(* Logix 5000 project; controller R400_500_XLS vendor 1 type 14 code 216 rev 31.11; software revision 31.01; part 3 of 32 *)
(* tags used below, declared in another part *)
   Alarm : SINT;   // Wait 3 seconds
   Ashutdown : SINT;   // Not Used
   CURRENT_CYCLE : DINT;
   CycleUsageArraySize : DINT;   // Size of the Cycle Usage Array
   CycleUsageDefaultUserName : STRING;   // Default User Name
   CycleUsageDefaultValue : UDT_CYCLE_USAGE;
   CycleUsageFirstEmptyIndex : DINT;   // Cycle Usage Array First Empty Index
   CycleUsageIterator : DINT;
   CycleUsagePrintoutCycleStartedCount : STRING;
   CycleUsagePrintoutHeader : STRING;
   CycleUsagePrintoutMessage : STRING;
   CycleUsagePrintoutSeparator : STRING;
   CycleUsageSearchCurrentUser : BOOL;
   CycleUsageSearchFirstEmptyIndex : BOOL;
   DESCALER : SINT;
   DRYING : DINT;   // Drying id number
   DRYING_HEAT_SENSITIVE_SEL : DINT;   // Drying heat sensitive
   DRYING_MODE_SEL : DINT;   // Drying mode selector index
   DRYING_TEMP_C_SEL : DINT;   // Drying temperature index
   DRYING_TEMP_F_SEL : DINT;   // Drying temperature index
   DRYING_TEMP_HIGH : REAL;   // Smart drying high temperature set point
   DRYING_TEMP_LOW : REAL;   // Smart drying low temperature set point
   DRYING_TEMP_STANDARD_LOW : REAL;   // Regular drying low temperature set point
   DRYING_TIME_LONG : DINT;   // Smart drying time for heat sensitive mode (in minute)
   DRYING_TIME_MIN_NUM : DINT;   // Drying time (minutes) numeric input index
   DRYING_TIME_SEC_NUM : DINT;   // Drying time (seconds) numeric input index
   DRYING_TIME_SHORT : DINT;   // Smart drying time for heat regular mode (in minute)
   ENVIRO_CARE : SINT;
   EXTRA_CARE : SINT;
   FINALRINSE_1 : DINT;   // Final rinse 1 id number
   FINALRINSE_2 : DINT;   // Final rinse 2 id number
   FINALRINSE_3 : DINT;   // Final rinse 3 id number
   FINALRINSE_4 : DINT;   // Final rinse 4 id number
   FINALRINSE_5 : DINT;   // Final rinse 5 id number
   FINALRINSE_6 : DINT;   // Final rinse 6 id number
   FINALRINSE_7 : DINT;   // Final rinse 7 id number
   FINALRINSE_8 : DINT;   // Final rinse 8 id number
   FINALRINSE_9 : DINT;   // Final rinse 9 id number
   FRINSE_COND_SET_POINT_NUM : DINT;   // Final rinse conductivity set point numeric input index
   FRINSE_DRAIN_SEL : DINT;   // Final rinse drained selector's index
   FRINSE_HEATING_SEL : DINT;   // Final rinse heating selector's index
   FRINSE_MIN_NUMBER_NUM : DINT;   // Final rinse minimum number of final rinse numeric input index
   FRINSE_NUMBER_NUM : DINT;   // Final rinse number of final rinse numeric input index
   FRINSE_RECIRC_SEL : DINT;   // Final rinse recirculated selector's index
   FRINSE_TIME_MIN_NUM : DINT;   // Final rinse time (minutes) numeric input index
   FRINSE_TIME_SEC_NUM : DINT;   // Final rinse time (seconds) numeric input index
   FRINSE_TYPE_SEL : DINT;   // Final rinse type selector's index
   HighLimt : REAL;
   LowLimt : REAL;
   M : DINT[5];   // Memory Bits
   NON_RECIRCULATED_FINAL_RINSE_MINUTES : DINT;   // Number of minutes for the non recirculated final rinse
   NON_RECIRCULATED_FINAL_RINSE_SECONDS : DINT;   // Number of seconds for the non recirculated final rinse
   PLASTIC_CARE : SINT;
   PREWASH_1 : DINT;   // Pre-wash 1 id number
   PREWASH_2 : DINT;   // Pre-wash 2 id number
   PREWASH_3 : DINT;   // Pre-wash 3 id number
   PREWASH_4 : DINT;   // Pre-wash 4 id number
   RINSE_1 : DINT;   // Rinse 1 id number
   RINSE_2 : DINT;   // Rinse 2 id number
   RINSE_3 : DINT;   // Rinse 3 id number
   RINSE_4 : DINT;   // Rinse 4 id number
   RINSE_CARE : SINT;
   Run : DINT;
   sCRLF : STRING;
   Service : DINT[2];   // Unused Service Mode Memory Bit
   sPrntArray : STRING[300];   // Printer String Array
   sSpaceCharacter : STRING;   // Space Character
   STANDARD : SINT;
   String : STRING[50];   // String
   SUMP_HIGH_VOLUME_400 : REAL;   // High sump volume
   SUMP_HIGH_VOLUME_500 : REAL;
   SUMP_LOW_VOLUME_400 : REAL;   // Low sump volume
   SUMP_LOW_VOLUME_500 : REAL;
   Supervisor : DINT;
   Tmr : TIMER[107];
   USER_DEFINED_10 : SINT;
   USER_DEFINED_11 : SINT;
   USER_DEFINED_7 : SINT;
   USER_DEFINED_8 : SINT;
   USER_DEFINED_9 : SINT;
   VENTING : DINT;   // Venting id number
   WASH_1 : DINT;   // Wash 1 id number
   WASH_2 : DINT;   // Wash 2 id number
   WASH_3 : DINT;   // Wash 3 id number
   WASH_4 : DINT;   // Wash 4 id number
   WASH_5 : DINT;   // Wash 5 id number
   WSH41_End_signal : BOOL;   // End of cycle signal
   AlarmTrigger : INT;   // Triggers the alarm screen if different of 0
   bAuditTrailExportButton : BOOL;
   bCSVExportHandshake : BOOL;
   bCycleOrAbortInProcess : BOOL;
   bONSAuditExportTrigger : BOOL;
   bONSAuditTrailEndOfCycle : BOOL;
   bONSBatchReportFileLocation : BOOL;
   bONSManualFileTransfer : BOOL;
   bPushButtonTransferFilesFromSDToUSB : BOOL;
   bTransferFilesFromSDToUSB : BOOL;
   bTransferFilesFromSDToUSBHandshakeLoad : BOOL;
   Current_Screen : DINT;
   CurrentUser : STRING;   // Current User
   CycleUsage : UDT_CYCLE_USAGE[50];
   CycleUsageListSelectedIndex : DINT;   // Current index selected in CycleUsage list
   CycleUsagePrint : BOOL;   // Print Cycle Usage
   CycleUsageResetAllValues : BOOL;   // Reset All Cycle Usage of all user
   CycleUsageResetDate : DINT[7];
   CycleUsageResetSelectedUser : BOOL;   // Reset Cycle Usage for the selected user
   DateTime : DINT[7];
   DISABLE : BOOL;   // Disable bit
   EmailSMSInt : INT[8];   // Email & SMS Notification Integer
   ENABLE : BOOL;   // Enable bit
   FALSE : BOOL;   // Always false bit
   NumInput : UDT_NUMERIC_INPUT[65];   // Numeric input
   PrintIndex : DINT;
   sBatchReportCSVName : STRING;
   sBatchReportFolderPath : STRING;
   Screen_Ctrl : DINT;   // PLC Screen Request
   sCycleCounter : STRING;
   sCycleForFileName : STRING;
   sHyphen : STRING;
   SumpHeatAlmRate : REAL;
   sUnderscore : STRING;
   tAuditTrailRemoteClearHistory : TIMER;
   Tpb : DINT[11];
   TpbImage : DINT[11];
   TRUE : BOOL;   // Always true bit
   udtAuditTrail : UDT_AuditTrail;
   udtCSVDataLogBatchReport : UDT_CSVDataLog;
   udtCSVExport : UDT_CSVExport;
   Unit : Hrdwre;   // Unit Configuration
(* MainProgram, continued *)

ROUTINE Constants   (* structured text *)
// Constant parameters
   // Program constants
   
   // General use constants
   TRUE := 1;				// Permanent, always true bit
   FALSE := 0;				// Permanent, always false bit
   ENABLE := 1;			// Used to ENABLE a bloc function
   DISABLE := 0;			// Used to DISABLE a bloc function
   
   // Sump water volume/level
   SUMP_LOW_VOLUME_400 := 22;        // Sump low water volume in liter
   SUMP_HIGH_VOLUME_400 := 36;       // Sump high water volume in liter
   SUMP_LOW_VOLUME_500 := 28.4;        // Sump low water volume in liter
   SUMP_HIGH_VOLUME_500 := 47.3;       // Sump high water volume in liter
   
   //XLSV10  DGB  2018-09-06 : Adjusted Treatments Constants
   // Treatment constants
   PREWASH_1 := 1;         // Pre-wash 1 id number
   PREWASH_2 := 2;         // Pre-wash 2 id number
   PREWASH_3 := 3;         // Pre-wash 3 id number
   PREWASH_4 := 4;         // Pre-wash 4 id number
   WASH_1 := 5;            // Wash 1 id number
   WASH_2 := 6;            // Wash 2 id number
   WASH_3 := 7;            // Wash 3 id number
   WASH_4 := 8;            // Wash 4 id number
   WASH_5 := 9;            // Wash 5 id number
   RINSE_1 := 10;           // Rinse 1 id number
   RINSE_2 := 11;           // Rinse 2 id number
   RINSE_3 := 12;           // Rinse 3 id number
   RINSE_4 := 13;           // Rinse 4 id number
   FINALRINSE_1 := 14;      // Final rinse 1 id number
   FINALRINSE_2 := 15;     // Final rinse 2 id number
   FINALRINSE_3 := 16;     // Final rinse 3 id number
   FINALRINSE_4 := 17;     // Final rinse 4 id number
   FINALRINSE_5 := 18;     // Final rinse 5 id number
   FINALRINSE_6 := 19;     // Final rinse 6 id number
   FINALRINSE_7 := 20;     // Final rinse 7 id number
   FINALRINSE_8 := 21;     // Final rinse 8 id number
   FINALRINSE_9 := 22;     // Final rinse 9 id number
   DRYING := 23;           // Drying id number
   VENTING := 24;          // Venting id number
   
   // Drying temperature and time
   DRYING_TEMP_LOW := 82.2;   // Smart drying low temperature set point
   DRYING_TEMP_HIGH := 115.6; // Smart drying high temperature set point
   //XLSV10  DGB  2018-09-10 : Changed Regular Low Temperature
   DRYING_TEMP_STANDARD_LOW := 65; // Standard drying high temperature set point
   DRYING_TIME_SHORT := 10;    // Smart drying time for heat regular mode (in minute)
   DRYING_TIME_LONG := 20;     // Smart drying time for heat sensitive mode (in minute)
   
   // Cycle constants
   EXTRA_CARE       := 0;
   ENVIRO_CARE      := 1;
   PLASTIC_CARE     := 2;
   STANDARD         := 3;
   RINSE_CARE       := 4;
   DESCALER         := 5;
   USER_DEFINED_7   := 6;
   USER_DEFINED_8   := 7;
   USER_DEFINED_9   := 8;
   USER_DEFINED_10  := 9;
   USER_DEFINED_11  := 10;
   CURRENT_CYCLE    := 11;
   
   
   // Control lists selectors indexes for the treatement modification
   DRYING_MODE_SEL := 14;
   DRYING_TEMP_C_SEL := 15;
   DRYING_TEMP_F_SEL := 16;
   DRYING_HEAT_SENSITIVE_SEL := 17;
   FRINSE_HEATING_SEL := 18;
   FRINSE_DRAIN_SEL := 19;
   FRINSE_RECIRC_SEL := 20;
   FRINSE_TYPE_SEL := 21;
   
   // Numeric input indexes for the treatement modification
   
   DRYING_TIME_MIN_NUM := 11;
   DRYING_TIME_SEC_NUM := 12;
   FRINSE_TIME_MIN_NUM := 14;
   FRINSE_TIME_SEC_NUM := 15;
   FRINSE_NUMBER_NUM := 16;
   FRINSE_MIN_NUMBER_NUM := 17;
   FRINSE_COND_SET_POINT_NUM := 18;
   
   // Non-recirculated final rinse time
   NON_RECIRCULATED_FINAL_RINSE_MINUTES := 0;
   NON_RECIRCULATED_FINAL_RINSE_SECONDS := 10;
   
   // Sump Heating alarm rate
   SumpHeatAlmRate:= 1.0;
   
   // Pure Water Tank low and High heating limit evaluation steam heated unit
   HighLimt:=0.1;
   LowLimt:=0.0;
   
   
   
   
   
END_ROUTINE

ROUTINE CycleUsage   (* ladder *)
// This Routine contains logic to manage the cycle usage
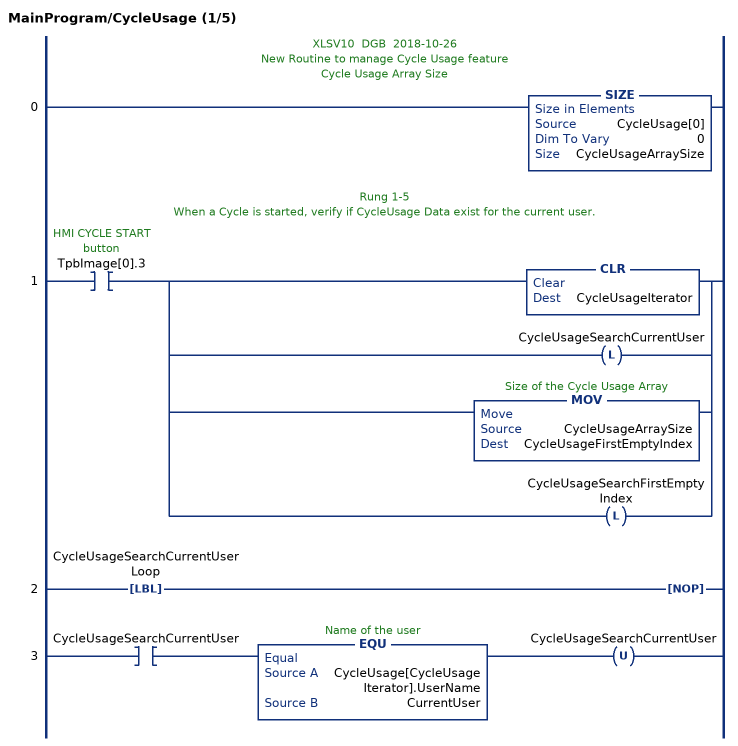
   // XLSV10  DGB  2018-10-26
   //  New Routine to manage Cycle Usage feature
   // Cycle Usage Array Size
   0: SIZE(CycleUsage[0],0,CycleUsageArraySize);
   // Rung 1-5
   // When a Cycle is started, verify if CycleUsage Data exist for the current user.
   1: XIC(TpbImage[0].3)[CLR(CycleUsageIterator) ,OTL(CycleUsageSearchCurrentUser) ,MOV(CycleUsageArraySize,CycleUsageFirstEmptyIndex) ,OTL(CycleUsageSearchFirstEmptyIndex) ];
   2: LBL(CycleUsageSearchCurrentUserLoop)NOP();
   3: XIC(CycleUsageSearchCurrentUser)EQU(CycleUsage[CycleUsageIterator].UserName,CurrentUser)OTU(CycleUsageSearchCurrentUser);
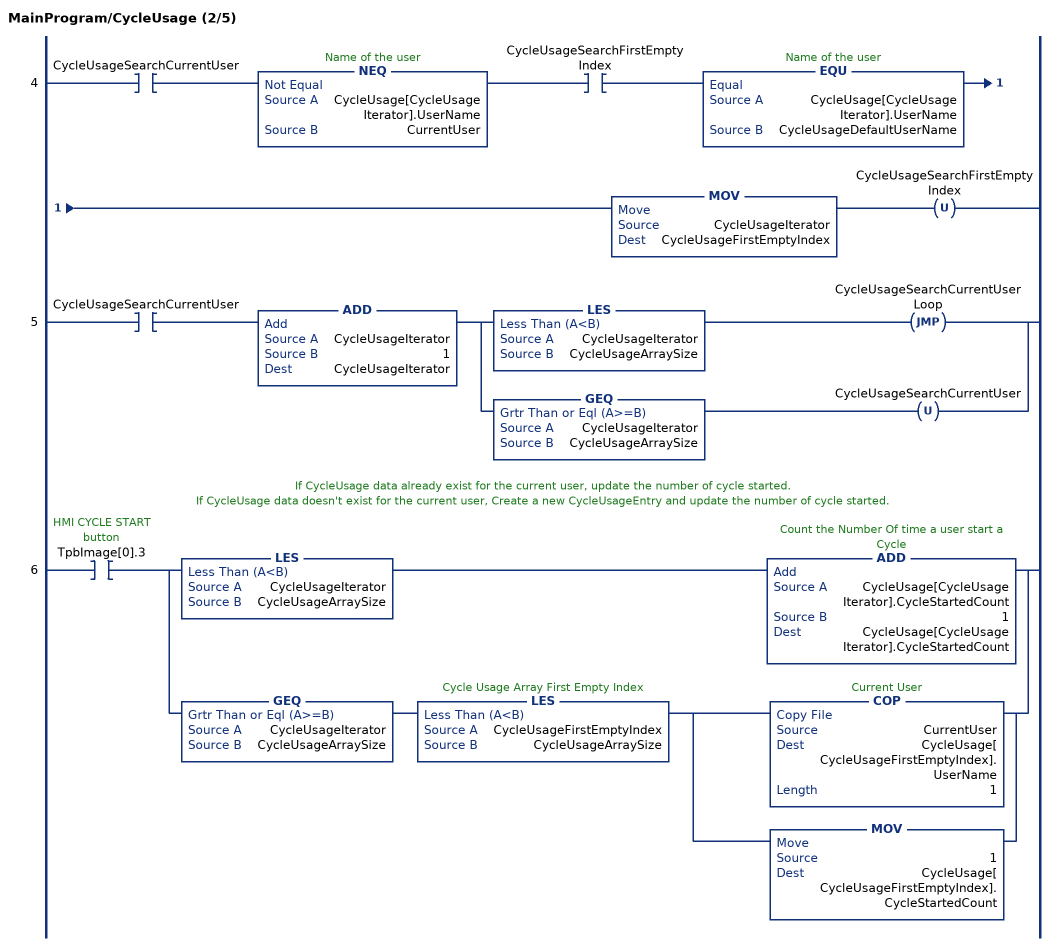
   4: XIC(CycleUsageSearchCurrentUser)NEQ(CycleUsage[CycleUsageIterator].UserName,CurrentUser)XIC(CycleUsageSearchFirstEmptyIndex)EQU(CycleUsage[CycleUsageIterator].UserName,CycleUsageDefaultUserName)MOV(CycleUsageIterator,CycleUsageFirstEmptyIndex)OTU(CycleUsageSearchFirstEmptyIndex);
   5: XIC(CycleUsageSearchCurrentUser)ADD(CycleUsageIterator,1,CycleUsageIterator)[LES(CycleUsageIterator,CycleUsageArraySize) JMP(CycleUsageSearchCurrentUserLoop) ,GEQ(CycleUsageIterator,CycleUsageArraySize) OTU(CycleUsageSearchCurrentUser) ];
   // If CycleUsage data already exist for the current user, update the number of cycle started.
   // If CycleUsage data doesn't exist for the current user, Create a new CycleUsageEntry and update the number of cycle started.
   6: XIC(TpbImage[0].3)[LES(CycleUsageIterator,CycleUsageArraySize) ADD(CycleUsage[CycleUsageIterator].CycleStartedCount,1,CycleUsage[CycleUsageIterator].CycleStartedCount) ,GEQ(CycleUsageIterator,CycleUsageArraySize) LES(CycleUsageFirstEmptyIndex,CycleUsageArraySize) [COP(CurrentUser,CycleUsage[CycleUsageFirstEmptyIndex].UserName,1) ,MOV(1,CycleUsage[CycleUsageFirstEmptyIndex].CycleStartedCount) ] ];
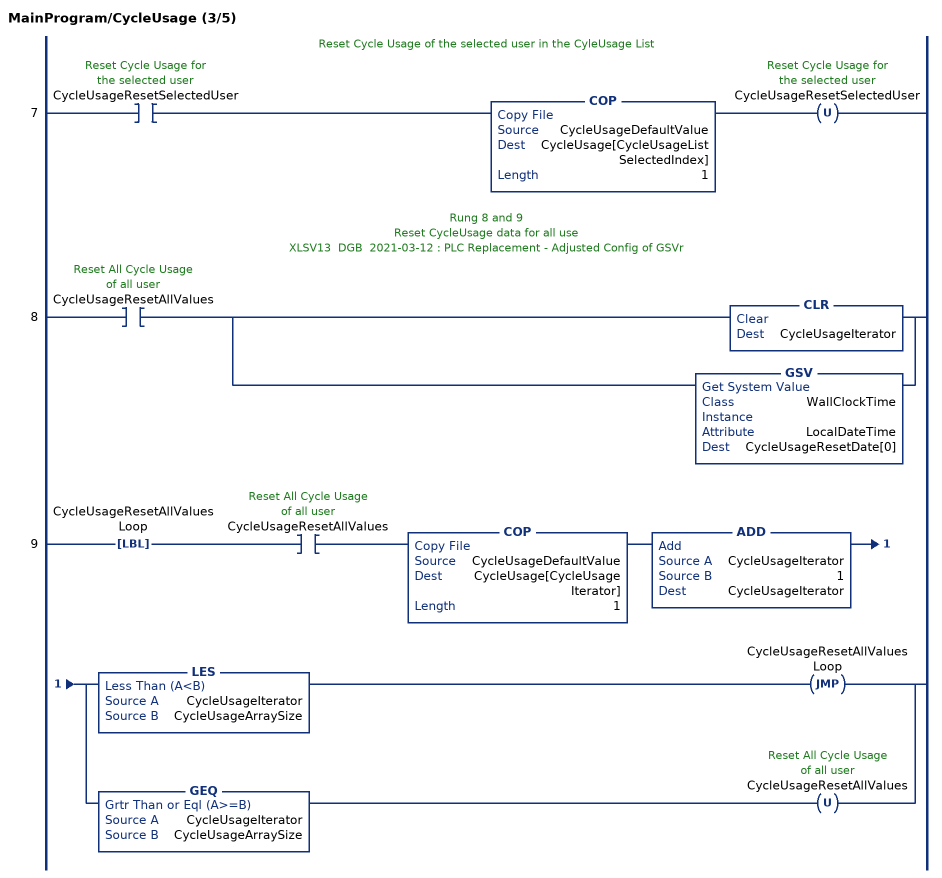
   // Reset Cycle Usage of the selected user in the CyleUsage List
   7: XIC(CycleUsageResetSelectedUser)COP(CycleUsageDefaultValue,CycleUsage[CycleUsageListSelectedIndex],1)OTU(CycleUsageResetSelectedUser);
   // Rung 8 and 9
   // Reset CycleUsage data for all use
   // XLSV13  DGB  2021-03-12 : PLC Replacement - Adjusted Config of GSVr
   8: XIC(CycleUsageResetAllValues)[CLR(CycleUsageIterator) ,GSV(WallClockTime,,LocalDateTime,CycleUsageResetDate[0]) ];
   9: LBL(CycleUsageResetAllValuesLoop)XIC(CycleUsageResetAllValues)COP(CycleUsageDefaultValue,CycleUsage[CycleUsageIterator],1)ADD(CycleUsageIterator,1,CycleUsageIterator)[LES(CycleUsageIterator,CycleUsageArraySize) JMP(CycleUsageResetAllValuesLoop) ,GEQ(CycleUsageIterator,CycleUsageArraySize) OTU(CycleUsageResetAllValues) ];
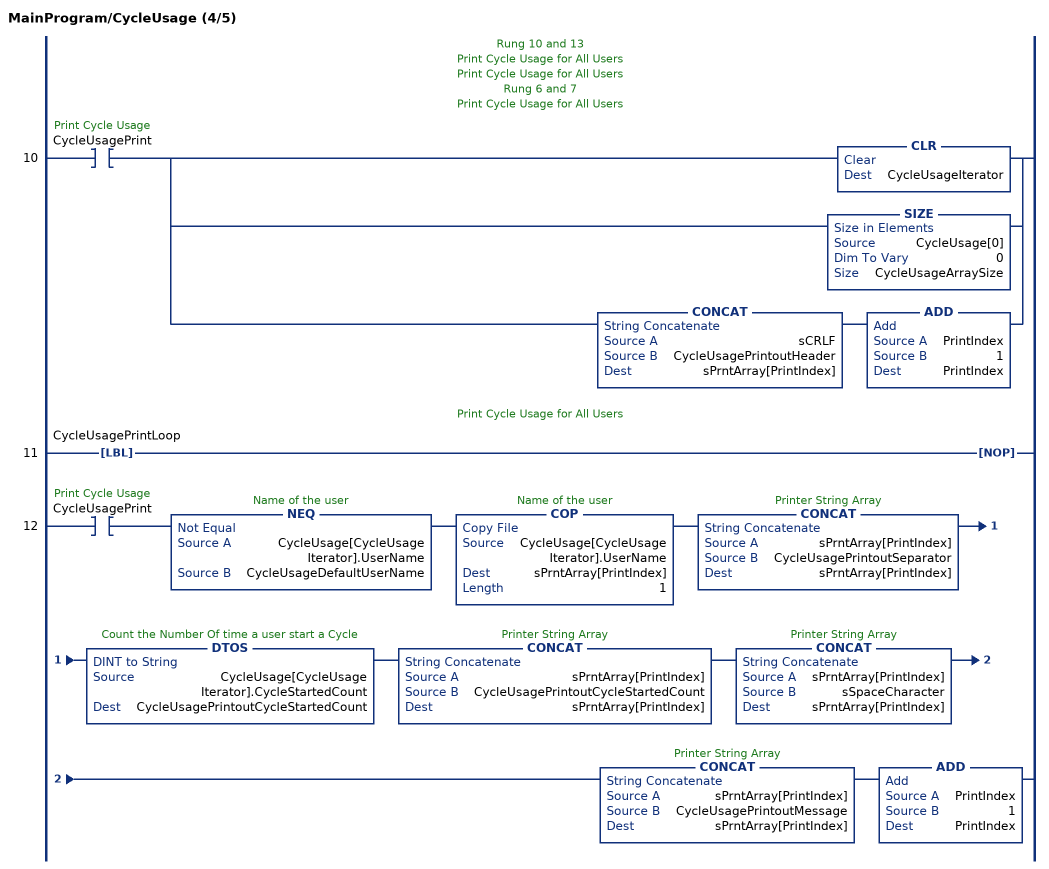
   // Rung 10 and 13
   //  Print Cycle Usage for All Users
   // Print Cycle Usage for All Users
   // Rung 6 and 7
   //  Print Cycle Usage for All Users
   10: XIC(CycleUsagePrint)[CLR(CycleUsageIterator) ,SIZE(CycleUsage[0],0,CycleUsageArraySize) ,CONCAT(sCRLF,CycleUsagePrintoutHeader,sPrntArray[PrintIndex]) ADD(PrintIndex,1,PrintIndex) ];
   // Print Cycle Usage for All Users
   11: LBL(CycleUsagePrintLoop)NOP();
   12: XIC(CycleUsagePrint)NEQ(CycleUsage[CycleUsageIterator].UserName,CycleUsageDefaultUserName)COP(CycleUsage[CycleUsageIterator].UserName,sPrntArray[PrintIndex],1)CONCAT(sPrntArray[PrintIndex],CycleUsagePrintoutSeparator,sPrntArray[PrintIndex])DTOS(CycleUsage[CycleUsageIterator].CycleStartedCount,CycleUsagePrintoutCycleStartedCount)CONCAT(sPrntArray[PrintIndex],CycleUsagePrintoutCycleStartedCount,sPrntArray[PrintIndex])CONCAT(sPrntArray[PrintIndex],sSpaceCharacter,sPrntArray[PrintIndex])CONCAT(sPrntArray[PrintIndex],CycleUsagePrintoutMessage,sPrntArray[PrintIndex])ADD(PrintIndex,1,PrintIndex);
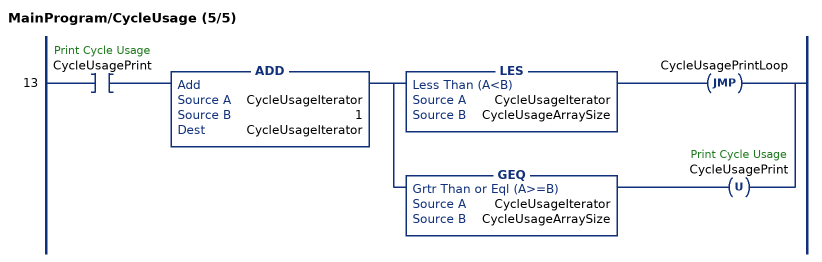
   13: XIC(CycleUsagePrint)ADD(CycleUsageIterator,1,CycleUsageIterator)[LES(CycleUsageIterator,CycleUsageArraySize) JMP(CycleUsagePrintLoop) ,GEQ(CycleUsageIterator,CycleUsageArraySize) OTU(CycleUsagePrint) ];
END_ROUTINE

ROUTINE EDS   (* ladder *)
// Manage Electronic Data Security Features
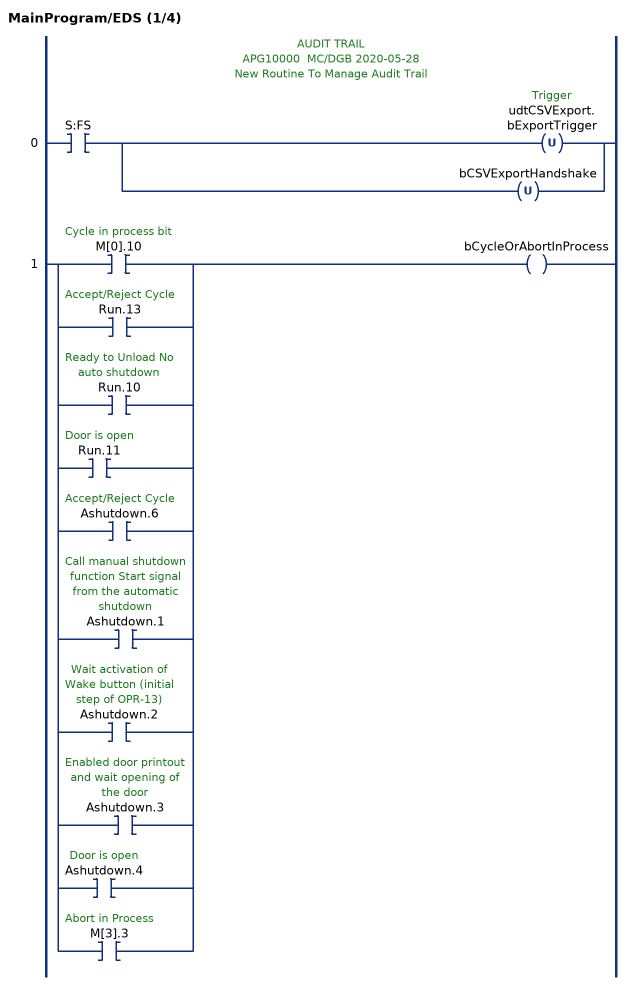
   // AUDIT TRAIL
   // APG10000  MC/DGB 2020-05-28
   // New Routine To Manage Audit Trail
   0: XIC(S:FS)[OTU(udtCSVExport.bExportTrigger) ,OTU(bCSVExportHandshake) ];
   1: [[XIC(M[0].10) ,[XIC(Run.13) ,XIC(Run.10) ,XIC(Run.11) ] ,[XIC(Ashutdown.6) ,XIC(Ashutdown.1) ,XIC(Ashutdown.2) ,XIC(Ashutdown.3) ,XIC(Ashutdown.4) ] ] ,XIC(M[3].3) ]OTE(bCycleOrAbortInProcess);
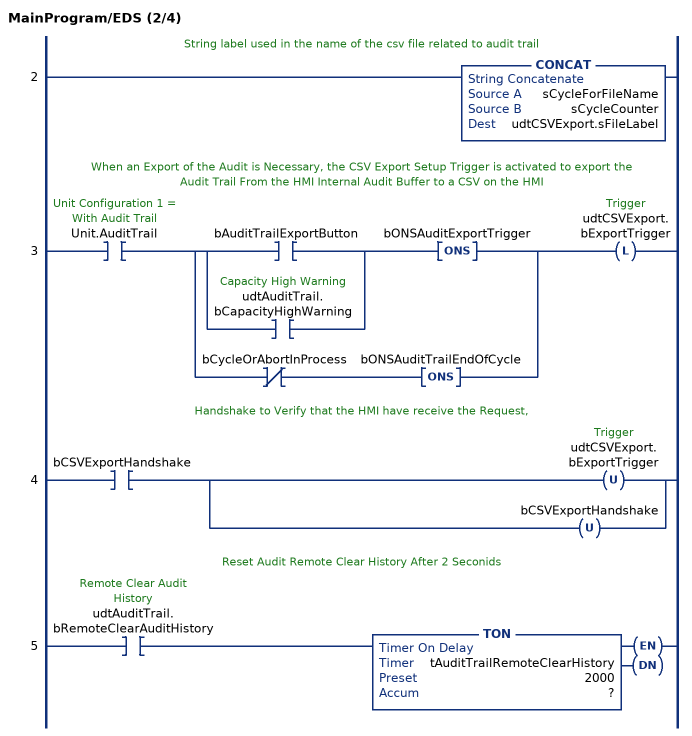
   // String label used in the name of the csv file related to audit trail
   2: CONCAT(sCycleForFileName,sCycleCounter,udtCSVExport.sFileLabel);
   // When an Export of the Audit is Necessary, the CSV Export Setup Trigger is activated to export the Audit Trail From the HMI Internal Audit Buffer to a CSV on the HMI
   3: XIC(Unit.AuditTrail)[[XIC(bAuditTrailExportButton) ,XIC(udtAuditTrail.bCapacityHighWarning) ] ONS(bONSAuditExportTrigger) ,XIO(bCycleOrAbortInProcess) ONS(bONSAuditTrailEndOfCycle) ]OTL(udtCSVExport.bExportTrigger);
   // Handshake to Verify that the HMI have receive the Request,
   4: XIC(bCSVExportHandshake)[OTU(udtCSVExport.bExportTrigger) ,OTU(bCSVExportHandshake) ];
   // Reset Audit Remote Clear History After 2 Seconids
   5: XIC(udtAuditTrail.bRemoteClearAuditHistory)TON(tAuditTrailRemoteClearHistory,?,?);
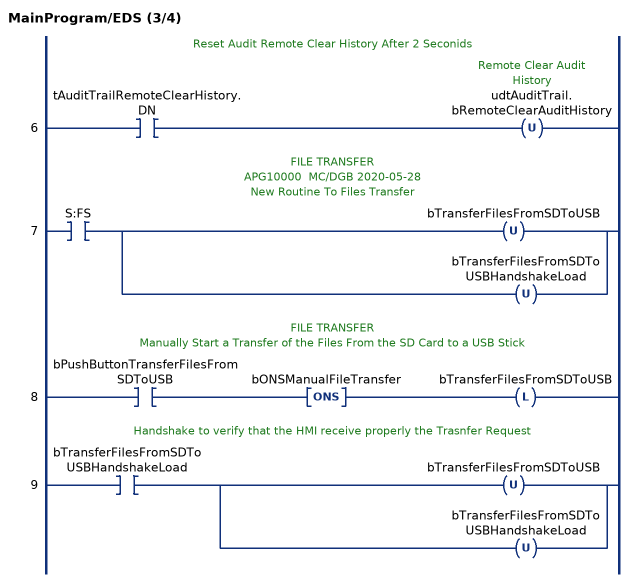
   // Reset Audit Remote Clear History After 2 Seconids
   6: XIC(tAuditTrailRemoteClearHistory.DN)OTU(udtAuditTrail.bRemoteClearAuditHistory);
   // FILE TRANSFER
   // APG10000  MC/DGB 2020-05-28
   // New Routine To Files Transfer
   7: XIC(S:FS)[OTU(bTransferFilesFromSDToUSB) ,OTU(bTransferFilesFromSDToUSBHandshakeLoad) ];
   // FILE TRANSFER
   // Manually Start a Transfer of the Files From the SD Card to a USB Stick
   8: XIC(bPushButtonTransferFilesFromSDToUSB)ONS(bONSManualFileTransfer)OTL(bTransferFilesFromSDToUSB);
   // Handshake to verify that the HMI receive properly the Trasnfer Request
   9: XIC(bTransferFilesFromSDToUSBHandshakeLoad)[OTU(bTransferFilesFromSDToUSB) ,OTU(bTransferFilesFromSDToUSBHandshakeLoad) ];
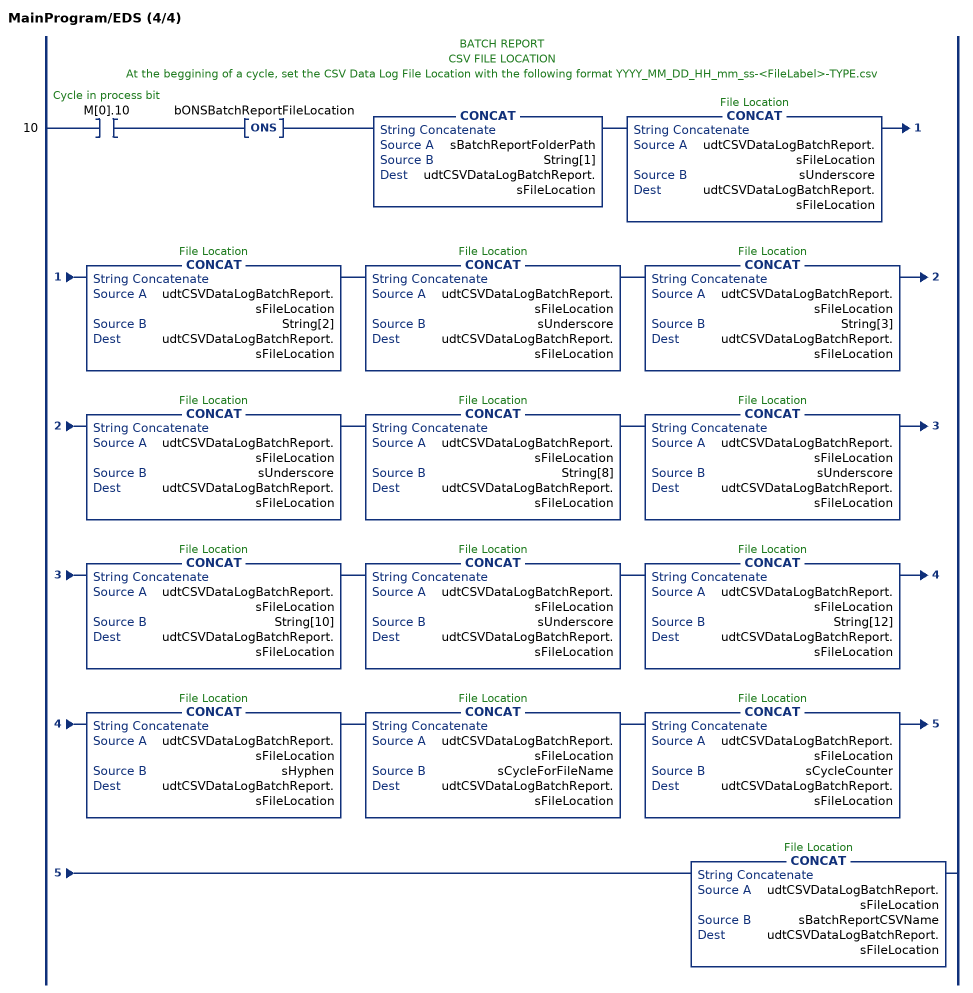
   // BATCH REPORT
   // CSV FILE LOCATION
   // At the beggining of a cycle, set the CSV Data Log File Location with the following format YYYY_MM_DD_HH_mm_ss-<FileLabel>-TYPE.csv
   10: XIC(M[0].10)ONS(bONSBatchReportFileLocation)CONCAT(sBatchReportFolderPath,String[1],udtCSVDataLogBatchReport.sFileLocation)CONCAT(udtCSVDataLogBatchReport.sFileLocation,sUnderscore,udtCSVDataLogBatchReport.sFileLocation)CONCAT(udtCSVDataLogBatchReport.sFileLocation,String[2],udtCSVDataLogBatchReport.sFileLocation)CONCAT(udtCSVDataLogBatchReport.sFileLocation,sUnderscore,udtCSVDataLogBatchReport.sFileLocation)CONCAT(udtCSVDataLogBatchReport.sFileLocation,String[3],udtCSVDataLogBatchReport.sFileLocation)CONCAT(udtCSVDataLogBatchReport.sFileLocation,sUnderscore,udtCSVDataLogBatchReport.sFileLocation)CONCAT(udtCSVDataLogBatchReport.sFileLocation,String[8],udtCSVDataLogBatchReport.sFileLocation)CONCAT(udtCSVDataLogBatchReport.sFileLocation,sUnderscore,udtCSVDataLogBatchReport.sFileLocation)CONCAT(udtCSVDataLogBatchReport.sFileLocation,String[10],udtCSVDataLogBatchReport.sFileLocation)CONCAT(udtCSVDataLogBatchReport.sFileLocation,sUnderscore,udtCSVDataLogBatchReport.sFileLocation)CONCAT(udtCSVDataLogBatchReport.sFileLocation,String[12],udtCSVDataLogBatchReport.sFileLocation)CONCAT(udtCSVDataLogBatchReport.sFileLocation,sHyphen,udtCSVDataLogBatchReport.sFileLocation)CONCAT(udtCSVDataLogBatchReport.sFileLocation,sCycleForFileName,udtCSVDataLogBatchReport.sFileLocation)CONCAT(udtCSVDataLogBatchReport.sFileLocation,sCycleCounter,udtCSVDataLogBatchReport.sFileLocation)CONCAT(udtCSVDataLogBatchReport.sFileLocation,sBatchReportCSVName,udtCSVDataLogBatchReport.sFileLocation);
END_ROUTINE

ROUTINE EMAIL_COMMAND   (* ladder *)
// EMAIL COMMAND, defines the different messages type
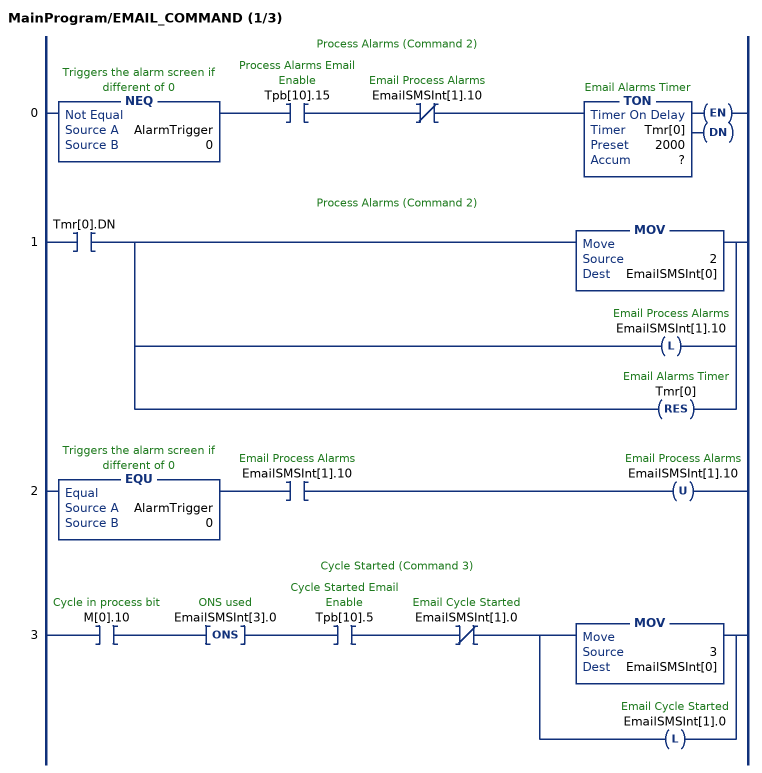
   // Process Alarms (Command 2)
   0: NEQ(AlarmTrigger,0)XIC(Tpb[10].15)XIO(EmailSMSInt[1].10)TON(Tmr[0],?,?);
   // Process Alarms (Command 2)
   1: XIC(Tmr[0].DN)[MOV(2,EmailSMSInt[0]) ,OTL(EmailSMSInt[1].10) ,RES(Tmr[0]) ];
   2: EQU(AlarmTrigger,0)XIC(EmailSMSInt[1].10)OTU(EmailSMSInt[1].10);
   // Cycle Started (Command 3)
   3: XIC(M[0].10)ONS(EmailSMSInt[3].0)XIC(Tpb[10].5)XIO(EmailSMSInt[1].0)[MOV(3,EmailSMSInt[0]) ,OTL(EmailSMSInt[1].0) ];
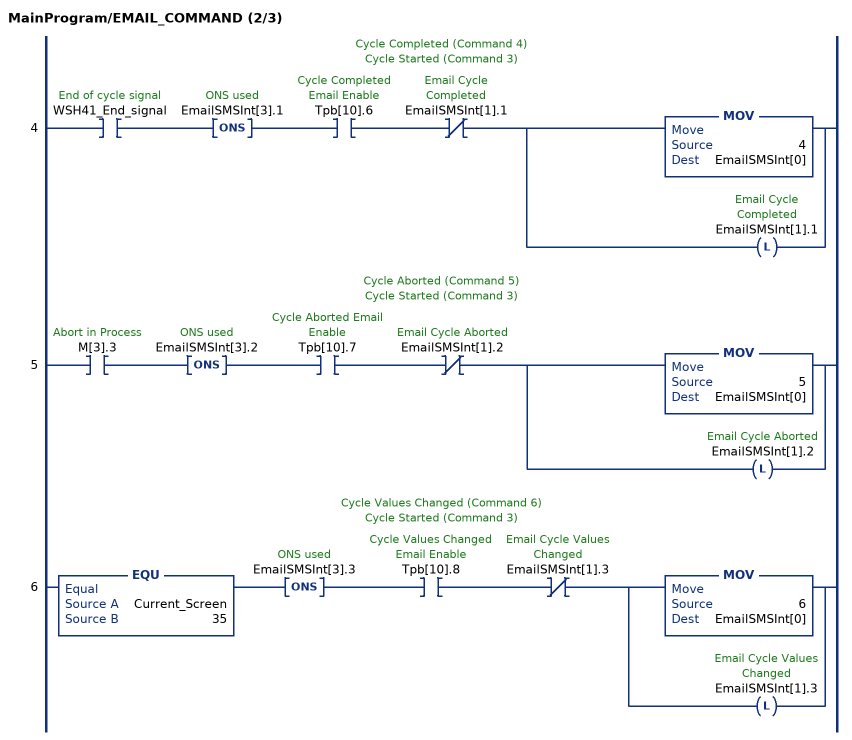
   // Cycle Completed (Command 4)
   // Cycle Started (Command 3)
   4: XIC(WSH41_End_signal)ONS(EmailSMSInt[3].1)XIC(Tpb[10].6)XIO(EmailSMSInt[1].1)[MOV(4,EmailSMSInt[0]) ,OTL(EmailSMSInt[1].1) ];
   // Cycle Aborted (Command 5)
   // Cycle Started (Command 3)
   5: XIC(M[3].3)ONS(EmailSMSInt[3].2)XIC(Tpb[10].7)XIO(EmailSMSInt[1].2)[MOV(5,EmailSMSInt[0]) ,OTL(EmailSMSInt[1].2) ];
   // Cycle Values Changed (Command 6)
   // Cycle Started (Command 3)
   6: EQU(Current_Screen,35)ONS(EmailSMSInt[3].3)XIC(Tpb[10].8)XIO(EmailSMSInt[1].3)[MOV(6,EmailSMSInt[0]) ,OTL(EmailSMSInt[1].3) ];
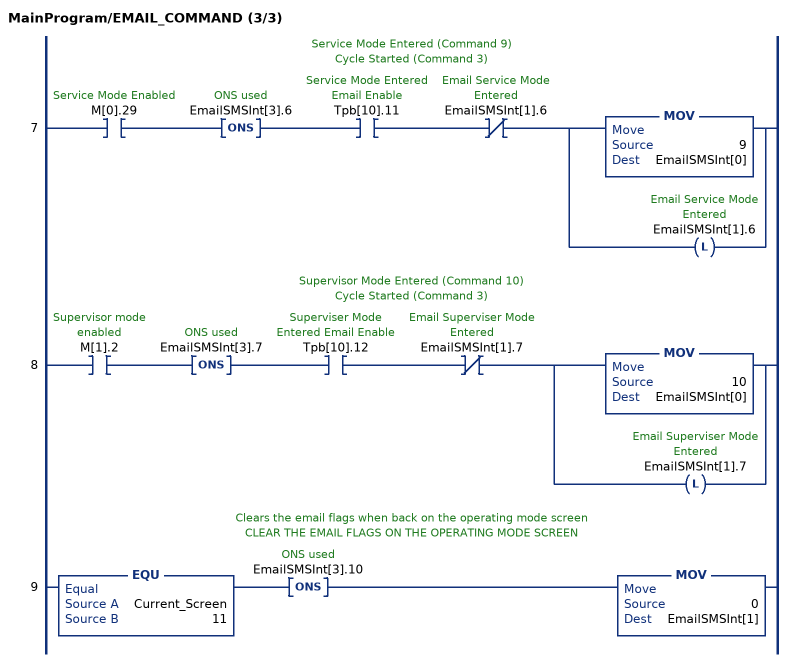
   // Service Mode Entered (Command 9)
   // Cycle Started (Command 3)
   7: XIC(M[0].29)ONS(EmailSMSInt[3].6)XIC(Tpb[10].11)XIO(EmailSMSInt[1].6)[MOV(9,EmailSMSInt[0]) ,OTL(EmailSMSInt[1].6) ];
   // Supervisor Mode Entered (Command 10)
   // Cycle Started (Command 3)
   8: XIC(M[1].2)ONS(EmailSMSInt[3].7)XIC(Tpb[10].12)XIO(EmailSMSInt[1].7)[MOV(10,EmailSMSInt[0]) ,OTL(EmailSMSInt[1].7) ];
   // Clears the email flags when back on the operating mode screen
   // CLEAR THE EMAIL FLAGS ON THE OPERATING MODE SCREEN
   9: EQU(Current_Screen,11)ONS(EmailSMSInt[3].10)MOV(0,EmailSMSInt[1]);
END_ROUTINE

ROUTINE EMAIL_PMPACK   (* ladder *)
// PREVENTIVE MAINTENANCE counters and triggers
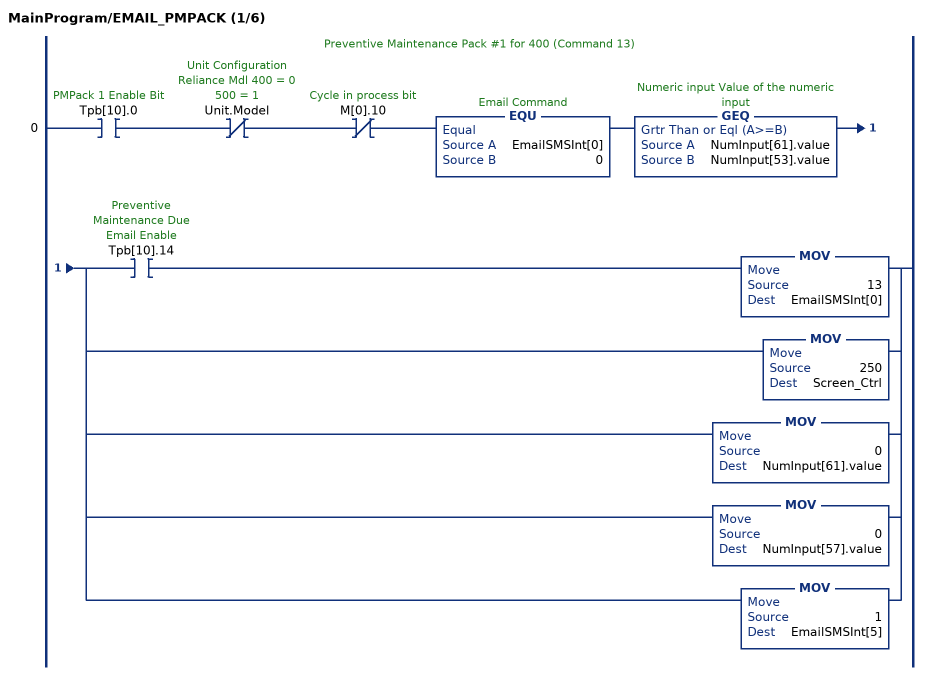
   // Preventive Maintenance Pack #1 for 400 (Command 13)
   0: XIC(Tpb[10].0)XIO(Unit.Model)XIO(M[0].10)EQU(EmailSMSInt[0],0)GEQ(NumInput[61].value,NumInput[53].value)[XIC(Tpb[10].14) MOV(13,EmailSMSInt[0]) ,MOV(250,Screen_Ctrl) ,MOV(0,NumInput[61].value) ,MOV(0,NumInput[57].value) ,MOV(1,EmailSMSInt[5]) ];
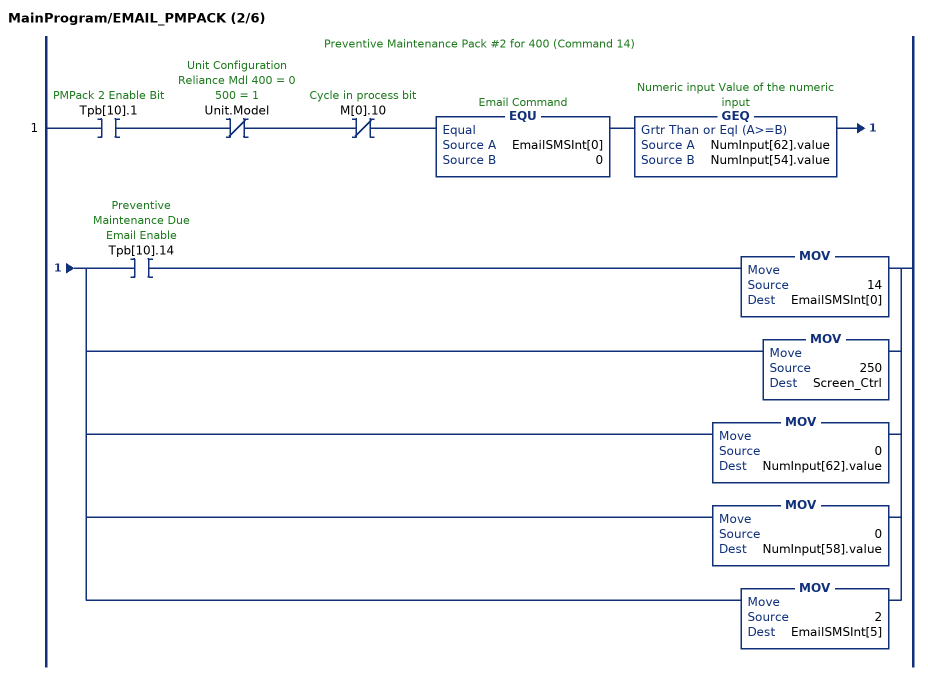
   // Preventive Maintenance Pack #2 for 400 (Command 14)
   1: XIC(Tpb[10].1)XIO(Unit.Model)XIO(M[0].10)EQU(EmailSMSInt[0],0)GEQ(NumInput[62].value,NumInput[54].value)[XIC(Tpb[10].14) MOV(14,EmailSMSInt[0]) ,MOV(250,Screen_Ctrl) ,MOV(0,NumInput[62].value) ,MOV(0,NumInput[58].value) ,MOV(2,EmailSMSInt[5]) ];
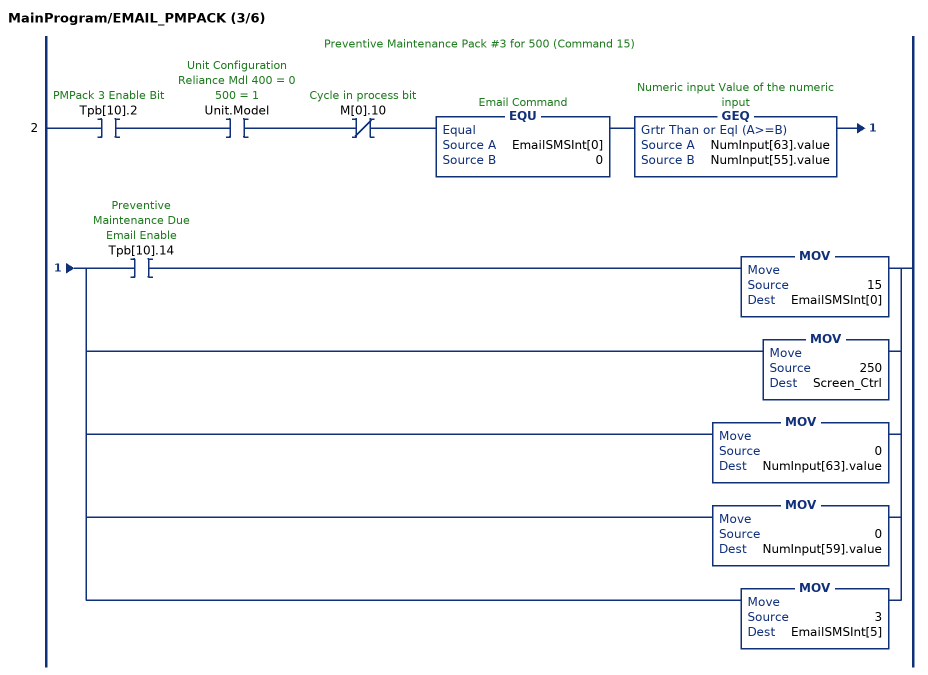
   // Preventive Maintenance Pack #3 for 500 (Command 15)
   2: XIC(Tpb[10].2)XIC(Unit.Model)XIO(M[0].10)EQU(EmailSMSInt[0],0)GEQ(NumInput[63].value,NumInput[55].value)[XIC(Tpb[10].14) MOV(15,EmailSMSInt[0]) ,MOV(250,Screen_Ctrl) ,MOV(0,NumInput[63].value) ,MOV(0,NumInput[59].value) ,MOV(3,EmailSMSInt[5]) ];
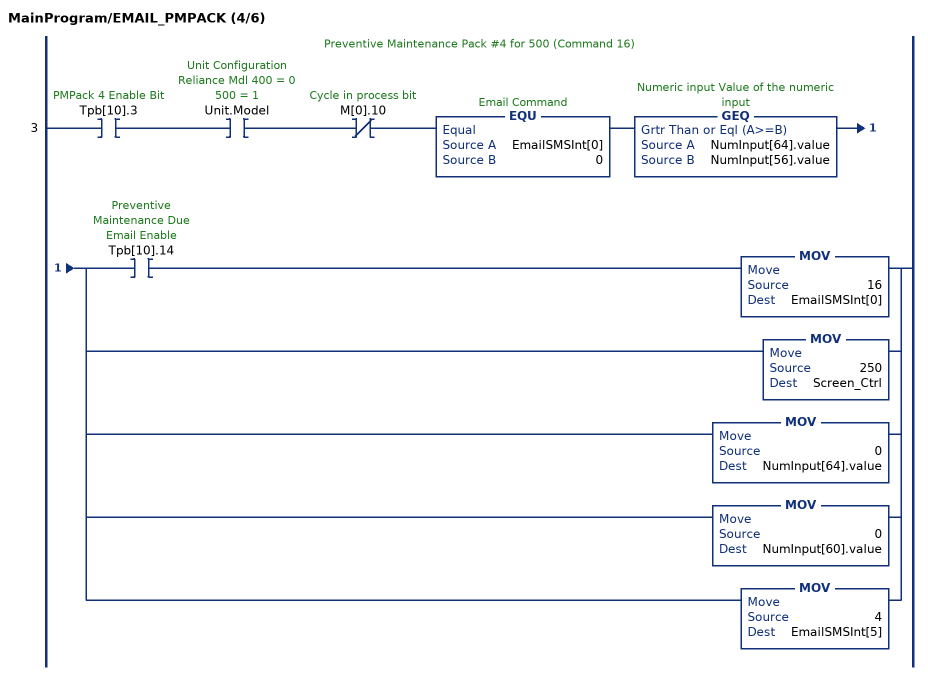
   // Preventive Maintenance Pack #4 for 500 (Command 16)
   3: XIC(Tpb[10].3)XIC(Unit.Model)XIO(M[0].10)EQU(EmailSMSInt[0],0)GEQ(NumInput[64].value,NumInput[56].value)[XIC(Tpb[10].14) MOV(16,EmailSMSInt[0]) ,MOV(250,Screen_Ctrl) ,MOV(0,NumInput[64].value) ,MOV(0,NumInput[60].value) ,MOV(4,EmailSMSInt[5]) ];
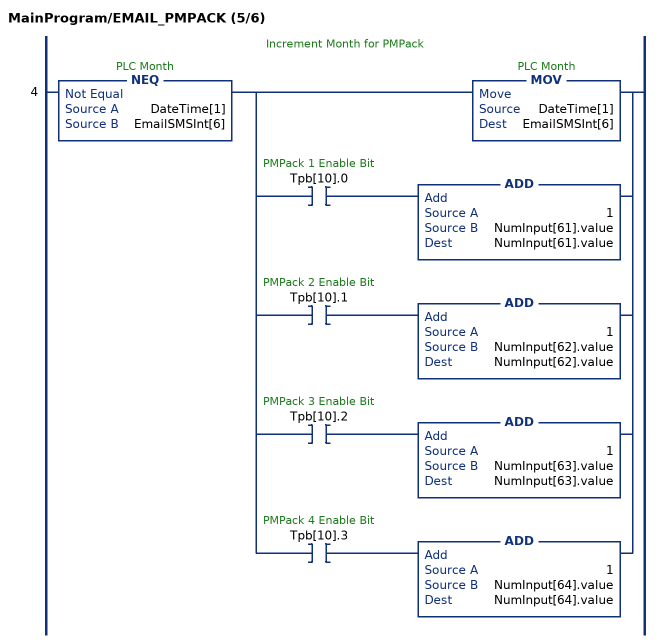
   // Increment Month for PMPack
   4: NEQ(DateTime[1],EmailSMSInt[6])[MOV(DateTime[1],EmailSMSInt[6]) ,XIC(Tpb[10].0) ADD(1,NumInput[61].value,NumInput[61].value) ,XIC(Tpb[10].1) ADD(1,NumInput[62].value,NumInput[62].value) ,XIC(Tpb[10].2) ADD(1,NumInput[63].value,NumInput[63].value) ,XIC(Tpb[10].3) ADD(1,NumInput[64].value,NumInput[64].value) ];
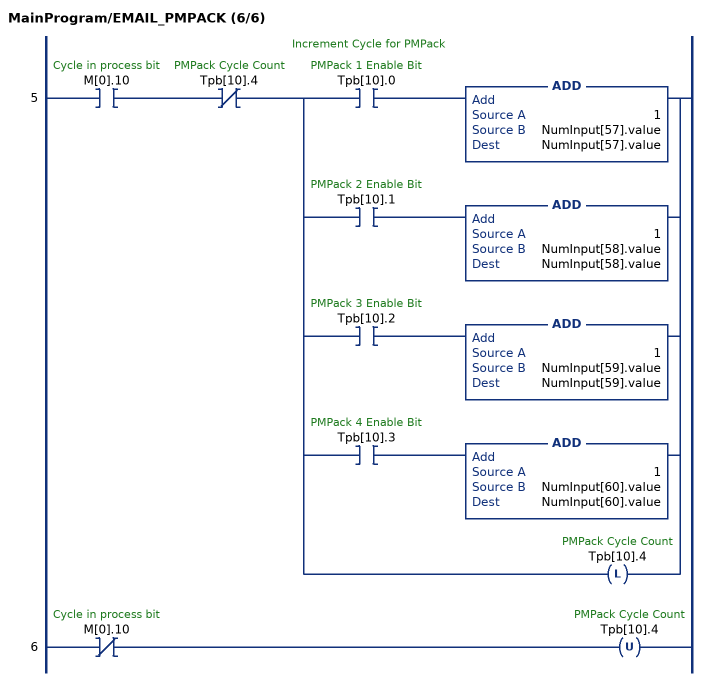
   // Increment Cycle for PMPack
   5: XIC(M[0].10)XIO(Tpb[10].4)[XIC(Tpb[10].0) ADD(1,NumInput[57].value,NumInput[57].value) ,XIC(Tpb[10].1) ADD(1,NumInput[58].value,NumInput[58].value) ,XIC(Tpb[10].2) ADD(1,NumInput[59].value,NumInput[59].value) ,XIC(Tpb[10].3) ADD(1,NumInput[60].value,NumInput[60].value) ,OTL(Tpb[10].4) ];
   6: XIO(M[0].10)OTU(Tpb[10].4);
END_ROUTINE
